# EPICS substitutions: db/user.substitutions
# SPDX-FileCopyrightText: 2006 Argonne National Laboratory
#
# SPDX-License-Identifier: EPICS

# Example substitutions file

file "db/circle.db" {
    { user = "RPI3" }
}

file "db/dbExample1.db" {
    { user = "RPI3" }
}

file db/dbExample2.db {
    pattern { user, no, scan }
        { "RPI3", 1, "1 second" }
        { "RPI3", 2, "2 second" }
        { "RPI3", 3, "5 second" }
}
